(* IEC 61131-3 sources: llm-plc-st-eval/data/processed_definitivo/gemini-3.1-pro-preview/I6/zero_shot, 3 files *)

(* ---- ejec_1.st ---- *)
FUNCTION_BLOCK FB_Temperatura
VAR_INPUT
    rawTemp : INT; // Señal analógica cruda del sensor (0 a 27648)
END_VAR

VAR_OUTPUT
    tempC : REAL; // Temperatura escalada en grados Celsius (0.0 a 100.0)
    enfriador : BOOL; // Comando de activación del enfriador
    almSensor : BOOL; // Alarma de sensor fuera de rango
END_VAR

// 1. Acondicionamiento y escalado de la señal
// Se convierte el valor entero a real y se escala al rango 0.0 - 100.0
tempC := (INT_TO_REAL(rawTemp) / 27648.0) * 100.0;

// 2. Detección de fallas del sensor (fuera de rango)
IF rawTemp < 0 OR rawTemp > 27648 THEN
    almSensor := TRUE;
ELSE
    almSensor := FALSE;
END_IF;

// 3. Control del enfriador con histéresis y seguridad
IF almSensor THEN
    // Por seguridad, si el sensor falla, se desactiva el enfriador
    enfriador := FALSE;
ELSIF tempC >= 80.0 THEN
    // Activar enfriador si alcanza o supera el umbral superior
    enfriador := TRUE;
ELSIF tempC <= 75.0 THEN
    // Desactivar enfriador si desciende al umbral inferior o menos
    enfriador := FALSE;
END_IF;
// Nota: Si tempC está entre 75.0 y 80.0, no se ejecuta ninguna condición,
// por lo que 'enfriador' conserva su estado anterior (histéresis).

END_FUNCTION_BLOCK

(* ---- ejec_2.st ---- *)
FUNCTION_BLOCK FB_Temperatura
VAR_INPUT
    rawTemp : INT; // Señal analógica cruda (0 a 27648)
END_VAR

VAR_OUTPUT
    tempC : REAL; // Temperatura escalada en grados Celsius (0.0 a 100.0)
    enfriador : BOOL; // Comando de activación del enfriador
    almSensor : BOOL; // Alarma de falla o fuera de rango del sensor
END_VAR

(* 1. Evaluación de alarma por señal fuera de rango *)
IF rawTemp < 0 OR rawTemp > 27648 THEN
    almSensor := TRUE;
ELSE
    almSensor := FALSE;
END_IF;

(* 2. Acondicionamiento y escalado de la señal a grados Celsius *)
tempC := (INT_TO_REAL(rawTemp) / 27648.0) * 100.0;

(* 3. Control del enfriador con histéresis y protección por alarma *)
IF almSensor THEN
    enfriador := FALSE; // Desactiva el enfriador por seguridad si hay falla
ELSIF tempC >= 80.0 THEN
    enfriador := TRUE;  // Activa el enfriador en el umbral superior
ELSIF tempC <= 75.0 THEN
    enfriador := FALSE; // Desactiva el enfriador en el umbral inferior
END_IF;
(* Nota: Si tempC está entre > 75.0 y < 80.0, la variable 'enfriador'
   no se reasigna, conservando así su estado actual (histéresis). *)

END_FUNCTION_BLOCK

(* ---- ejec_3.st ---- *)
FUNCTION_BLOCK FB_Temperatura
VAR_INPUT
    rawTemp : INT; // Señal analógica cruda (0 a 27648)
END_VAR

VAR_OUTPUT
    tempC : REAL; // Temperatura escalada en grados Celsius (0.0 a 100.0)
    enfriador : BOOL; // Estado del enfriador
    almSensor : BOOL; // Alarma de sensor fuera de rango
END_VAR

// 1. Evaluación de alarma por fuera de rango
IF rawTemp < 0 OR rawTemp > 27648 THEN
    almSensor := TRUE;
ELSE
    almSensor := FALSE;
END_IF;

// 2. Acondicionamiento y escalado de la señal a REAL (0.0 - 100.0)
tempC := (INT_TO_REAL(rawTemp) / 27648.0) * 100.0;

// 3. Control del enfriador con histéresis y enclavamiento por alarma
IF almSensor THEN
    // Por seguridad, si el sensor falla, se desactiva el enfriador
    enfriador := FALSE;
ELSE
    // Lógica de histéresis
    IF tempC >= 80.0 THEN
        enfriador := TRUE;
    ELSIF tempC <= 75.0 THEN
        enfriador := FALSE;
    END_IF;
    // Si tempC está entre 75.0 y 80.0, 'enfriador' conserva su estado anterior
END_IF;

END_FUNCTION_BLOCK
